Staubli VAL3: physicalIO.pgx

program physicalIO()
// Suction tool inputs and outputs
begin
  // Only the suction tool is controlled in Levels 1 and 2.
  while true
    partOnTool = io:bIn0 == true
    io:bOut0 = vacuumOn
    io:bOut1 = blowOn
    ioReady = true
    delay(0.01)
  endWhile
end
